(* IEC 61131-3 sources: kns-pump-station/tests/POUs/Station/FB_Annunciator_Test, 10 files *)

(* ---- HornOffWhenAllAcked.method.decl.st ---- *)
// 04 §14: квитирование всех High/Critical выключает сирену
METHOD PRIVATE HornOffWhenAllAcked
VAR
    fbDut  : FB_Annunciator;            // ФБ под тестом
    fbTime : PL.FB_FakeTime;            // подменное время, старт 1 ч
END_VAR

(* ---- HornOnNewHighUnack.method.decl.st ---- *)
// 04 §14, PMI-36: новая неквитированная High/Critical (рост udiNewHighSeq) включает сирену; первый вызов принимает
// счётчик как есть
METHOD PRIVATE HornOnNewHighUnack
VAR
    fbDut  : FB_Annunciator;            // ФБ под тестом
    fbTime : PL.FB_FakeTime;            // подменное время, старт 1 ч
END_VAR

(* ---- K1DeenergizedOnActiveHigh.method.decl.st ---- *)
// 04 §14, PMI-17, PMI-20: K1 под напряжением в норме, обесточено при активной High или Critical; Medium — нет
METHOD PRIVATE K1DeenergizedOnActiveHigh
VAR
    fbDut  : FB_Annunciator;            // ФБ под тестом
    fbTime : PL.FB_FakeTime;            // подменное время, старт 1 ч
END_VAR

(* ---- LampBlinksAt1Hz.method.decl.st ---- *)
// 04 §14, PMI-36: HL1 мигает 1 Гц при неквитированных Medium и выше — 0,5 с горит, 0,5 с нет; Low не мигает
METHOD PRIVATE LampBlinksAt1Hz
VAR
    fbDut  : FB_Annunciator;            // ФБ под тестом
    fbTime : PL.FB_FakeTime;            // подменное время, старт 1 ч
    uiStep : UINT;                    // шаг 100 мс
    fbDut2 : FB_Annunciator;          // второй экземпляр: только Low
END_VAR

(* ---- LampBlinksAt1Hz.method.impl.st ---- *)
coUnit.TEST('Annunciator_LampBlinksAt1Hz_A14_PMI36');

fbDut.auiUnack[2] := 1;
fbDut(itfTime := fbTime);
AssertTrue(Condition := fbDut.xLamp, Message := 'on at blink start');
FOR uiStep := 1 TO 4 DO
    fbTime.Advance(tStep := T#100MS);
    fbDut(itfTime := fbTime);
END_FOR
AssertTrue(Condition := fbDut.xLamp, Message := 'on at 0.4 s');
fbTime.Advance(tStep := T#100MS);
fbDut(itfTime := fbTime);
AssertFalse(Condition := fbDut.xLamp, Message := 'off at 0.5 s');
FOR uiStep := 1 TO 4 DO
    fbTime.Advance(tStep := T#100MS);
    fbDut(itfTime := fbTime);
END_FOR
AssertFalse(Condition := fbDut.xLamp, Message := 'off at 0.9 s');
fbTime.Advance(tStep := T#100MS);
fbDut(itfTime := fbTime);
AssertTrue(Condition := fbDut.xLamp, Message := 'on again at 1.0 s');
fbDut2.auiUnack[1] := 1;
fbDut2(itfTime := fbTime);
AssertFalse(Condition := fbDut2.xLamp OR fbDut2.xHorn, Message := 'Low only: no lamp, no horn');

coUnit.TEST_FINISHED();

(* ---- LampSteadyWhenActiveAcked.method.decl.st ---- *)
// 04 §14, PMI-36 шаг 3: активные квитированные — HL1 горит постоянно; нет активных — погашена
METHOD PRIVATE LampSteadyWhenActiveAcked
VAR
    fbDut  : FB_Annunciator;            // ФБ под тестом
    fbTime : PL.FB_FakeTime;            // подменное время, старт 1 ч
    uiStep : UINT;                    // шаг 100 мс
    xEverOff : BOOL;                  // лампа гасла
END_VAR

(* ---- LampSteadyWhenActiveAcked.method.impl.st ---- *)
coUnit.TEST('Annunciator_LampSteadyWhenActiveAcked_A14_PMI36');

fbDut.auiActive[2] := 1;
fbDut(itfTime := fbTime);
FOR uiStep := 1 TO 20 DO
    fbTime.Advance(tStep := T#100MS);
    fbDut(itfTime := fbTime);
    xEverOff := xEverOff OR NOT fbDut.xLamp;
END_FOR
AssertFalse(Condition := xEverOff, Message := 'steady on while active acked');
fbDut.auiActive[2] := 0;
fbDut(itfTime := fbTime);
AssertFalse(Condition := fbDut.xLamp, Message := 'off without alarms');

coUnit.TEST_FINISHED();

(* ---- SilenceStopsHornUntilNextNew.method.decl.st ---- *)
// 04 §14, PMI-36 шаг 2: «Звук» выключает сирену до следующей новой тревоги
METHOD PRIVATE SilenceStopsHornUntilNextNew
VAR
    fbDut  : FB_Annunciator;            // ФБ под тестом
    fbTime : PL.FB_FakeTime;            // подменное время, старт 1 ч
END_VAR

(* ---- TimeBackwardsRestartsBlink.method.decl.st ---- *)
// Время назад — мигание HL1 начинается заново с фазы «горит»
METHOD PRIVATE TimeBackwardsRestartsBlink
VAR
    fbDut  : FB_Annunciator;            // ФБ под тестом
    fbTime : PL.FB_FakeTime;            // подменное время, старт 1 ч
    uiStep : UINT;                    // шаг 100 мс
END_VAR

(* ---- TimeBackwardsRestartsBlink.method.impl.st ---- *)
coUnit.TEST('Annunciator_TimeBackwardsRestartsBlink_A14');

fbDut.auiUnack[2] := 1;
fbDut(itfTime := fbTime);
FOR uiStep := 1 TO 5 DO
    fbTime.Advance(tStep := T#100MS);
    fbDut(itfTime := fbTime);
END_FOR
AssertFalse(Condition := fbDut.xLamp, Message := 'off at 0.5 s');
fbTime.SetNow(ltValue := LTIME#59M);
fbDut(itfTime := fbTime);
AssertTrue(Condition := fbDut.xLamp, Message := 'blink restarted on time jump: on');
FOR uiStep := 1 TO 5 DO
    fbTime.Advance(tStep := T#100MS);
    fbDut(itfTime := fbTime);
END_FOR
AssertFalse(Condition := fbDut.xLamp, Message := 'off 0.5 s after restart');

coUnit.TEST_FINISHED();
